// TIA Portal V20 export
Screen "Pop-up_CURVE_STD-CYCLETIMES_Popup"  640x320
  ScreenItem "Background" at 0,0 size 640x320  Type=HmiRectangle
  ScreenItem "趋势控件_1" at 0,0 size 640x320  Type=HmiTrendControl
  ScreenItem "ButtonClose" at 568,0 size 72x32  Type=HmiButton
